RoboDK station: Senior Project 6612247056.rdk

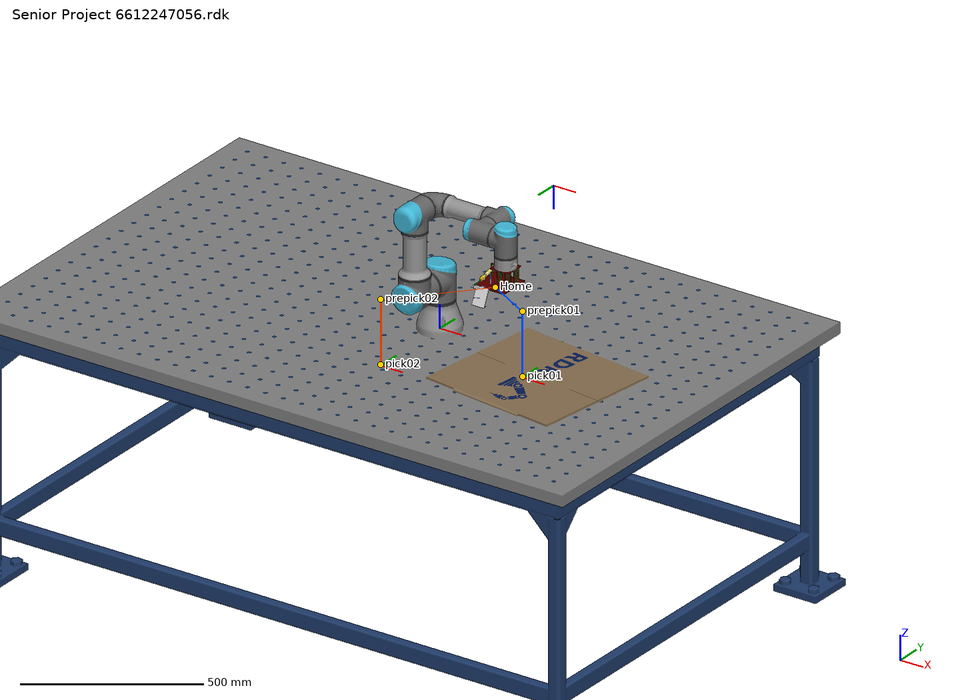
[picture v0: the station drawn from its stored meshes, robots at their saved joint values, targets as dots, program paths as lines]
Station Tast (saved by RoboDK 6.0.1). Poses are relative to the parent item; angles as X-Y-Z fixed-axis rotations.
  - frame Table at (0, 0, 0) mm
    - object Table at (-760, 0, 0) mm, size 2020 x 1340 x 800 mm, geometry from Table-2000x1200x800mm.sld
    - target Home (Cartesian target) at (261.4, -110.4, 243.15) mm, rotated rx -180 ry 0 rz -90 deg; joints [0, -90, -90, -90, 90, 0] of UR3
    - frame Camera 1 at (450, -100, 600) mm, rotated rx 180 ry 0 rz 0 deg
      - camera Camera 1
    - object BOX at (374.64, -51.63, 2) mm, rotated rx 0 ry 0.01 rz -7.34 deg, size 444 x 419.7 x 11.5 mm, geometry from Box-215x215mm-Unfolded.sld
  - frame UR3 Base at (0, 0, 0) mm
    - robot UR3: 6 axes, payload 3 kg, reach 500 mm, repeatability 0.1 mm, weight 11 kg
        modified DH rows (alpha deg, a mm, theta deg, d mm): 0, 0, 0, 151.9; 90, 0, 180, 0; 0, 243.65, 0, 0; 0, 213, 0, 110.4; -90, 0, 0, 83.4; 90, 0, 180, 82.4
        joint limits [-360, -360, -360, -360, -360, -360] to [360, 360, 360, 360, 360, 360]; home [0, -90, -90, 0, 90, 0]; saved at [0, -90, -90, -90, 90, 0]
      - tool Assem1, TCP at (0, 35, 70) mm, size 142.5 x 102 x 100.1 mm, geometry from Assem1.STEP
  - frame Orinal_Box at (360, -120, 0) mm
    - target prepick01 (Cartesian target) at (0, 0, 200) mm, rotated rx 180 ry 0 rz -90 deg; joints [20.517, -90.713, -100.969, -78.318, 90, 20.517] of UR3
    - target pick01 (Cartesian target) at (0, 0, 2) mm, rotated rx -180 ry 0 rz -90 deg; joints [-1.388, -136.982, -93.252, -39.765, 90.001, -1.388] of UR3
  - frame Orinal_Box(2) at (0, -280, 0) mm
    - target prepick02 (Cartesian target) at (0, 0, 200) mm, rotated rx -179.99 ry 0 rz 178.23 deg; joints [-68.924, -88.183, -103.474, -78.333, 90.001, 22.846] of UR3
    - target pick02 (Cartesian target) at (0, 0, 2) mm, rotated rx 179.99 ry 0 rz -179.49 deg; joints [-69.427, -124.075, -125.27, -20.665, 90, 20.063] of UR3
  - program Prog1 (1 instructions, listed below)
  - program pick (10 instructions, listed below)
  - program Place (8 instructions, listed below)
  - Python program Prog5 (listed below)
  - program Run (3 instructions, listed below)
  - Python program ur3_vision_pick_place (listed below)
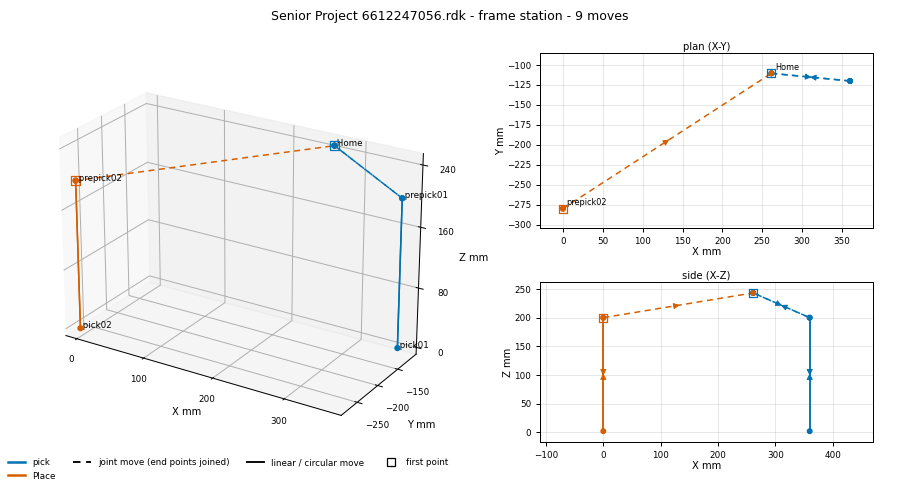
[picture p0: tool path of Senior Project 6612247056.rdk in frame station, 9 of 9 moves have a stored position in this frame; points joined in program order, loops and branches not executed]

--- program Prog1 (robot UR3) ---
  Move objects

--- program pick (robot UR3) ---
  ตั้งค่าRef: Table
  ตั้งค่าเครื่องมือ: Assem1
  MoveJ (Home)
  ตั้งค่าRef: Orinal_Box
  MoveJ (prepick01)
  MoveL (pick01)
  Attach to Assem1
  MoveL (prepick01)
  ตั้งค่าRef: Table
  MoveJ (Home)

--- program Place (robot UR3) ---
  ตั้งค่าRef: Orinal_Box(2)
  ตั้งค่าเครื่องมือ: Tool 1 at (0, 35, 70) mm
  MoveJ (prepick02)
  MoveL (pick02)
  ถอดออกจาก Assem1
  MoveL (prepick02)
  ตั้งค่าRef: Table
  MoveJ (Home)

--- Python program Prog5 ---
from robodk import robolink

RDK = robolink.Robolink()

# ดึงโปรแกรมมารันตรงๆ
prog_pick = RDK.Item('pick', robolink.ITEM_TYPE_PROGRAM)
prog_place = RDK.Item('Place', robolink.ITEM_TYPE_PROGRAM)

print("กำลังรันโปรแกรม Pick...")
prog_pick.RunProgram()


print("กำลังรันโปรแกรม Place...")
prog_place.RunProgram()

--- program Run (robot UR3) ---
  โทร Prog1
  โทร pick
  โทร Place

--- Python program ur3_vision_pick_place ---
"""
===============================================================================
UR3 Vision-Guided Pick & Place System with YOLOv8 & RoboDK
===============================================================================
Senior Project 6612247047
- YOLOv8 Model: Box_Logo.v2i.yolov8 (best (2).pt)
- RoboDK Station: Senior Project 6612247047 (UR3 Robot + Assem1 Gripper + BOX)
- Collision-Free Safe Execution via Home Posture
===============================================================================
"""

from robodk.robolink import *
from robodk.robomath import *
from ultralytics import YOLO
import cv2
import os
import time

# -----------------------------------------------------------------------------
# 1. Configuration & Initializations
# -----------------------------------------------------------------------------
MODEL_PATH = r'f:\New folder\best (2).pt'
SNAPSHOT_PATH = r'f:\New folder\temp_cam_snapshot.png'
ROBOT_SPEED = 80  # Speed in mm/s for safe motion

print("=" * 60)
print("  UR3 Vision-Guided Pick & Place System starting...")
print("=" * 60)

# Load YOLOv8 Model
if not os.path.exists(MODEL_PATH):
    raise FileNotFoundError(f"Model file not found at: {MODEL_PATH}")

print(f"[AI] Loading YOLOv8 model: {MODEL_PATH}...")
model = YOLO(MODEL_PATH)
print(f"[AI] Model classes loaded: {model.names}")

# Connect to RoboDK
print("[RoboDK] Connecting to RoboDK...")
RDK = Robolink()

if not RDK.Connect():
    print("[ERROR] Could not connect to RoboDK! Please ensure RoboDK is running.")
    exit(1)

station = RDK.ActiveStation()
print(f"[RoboDK] Connected to station: '{station.Name()}'")

# Get Items from RoboDK Station
robot = RDK.Item('UR3', ITEM_TYPE_ROBOT)
gripper = RDK.Item('Assem1', ITEM_TYPE_TOOL)
if not gripper.Valid():
    gripper = RDK.Item('gripper', ITEM_TYPE_TOOL)

target_item = RDK.Item('BOX', ITEM_TYPE_OBJECT)
if not target_item.Valid():
    target_item = RDK.Item('box', ITEM_TYPE_OBJECT)

home_target = RDK.Item('Home', ITEM_TYPE_TARGET)
prepick01 = RDK.Item('prepick01', ITEM_TYPE_TARGET)
pick01 = RDK.Item('pick01', ITEM_TYPE_TARGET)
prepick02 = RDK.Item('prepick02', ITEM_TYPE_TARGET)
pick02 = RDK.Item('pick02', ITEM_TYPE_TARGET)

table_frame = RDK.Item('Table', ITEM_TYPE_FRAME)
if not table_frame.Valid():
    table_frame = target_item.Parent()

cam_item = RDK.Item('Camera 1')

# Validate essential items
if not robot.Valid():
    print("[ERROR] Robot 'UR3' not found in RoboDK station!")
    exit(1)
if not target_item.Valid():
    print("[ERROR] Object 'BOX' not found in RoboDK station!")
    exit(1)

print("[RoboDK] All essential robot and station items loaded successfully.")

# Set safe robot speed
robot.setSpeed(ROBOT_SPEED)

# -----------------------------------------------------------------------------
# 2. Collision-Free Pick and Place Routine
# -----------------------------------------------------------------------------
def execute_safe_pick_and_place():
    """
    Executes a safe step-by-step pick and place operation for UR3:
    1. Move to Home (safe posture)
    2. Approach prepick01 (hover over source)
    3. Move to pick01 (pick position)
    4. Attach object BOX to gripper Assem1
    5. Retract up to prepick01
    6. Return to Home (safe transit posture avoiding self-collision)
    7. Move to prepick02 (hover over target destination)
    8. Move to pick02 (place position)
    9. Detach object BOX to table frame
    10. Retract up to prepick02
    11. Return safely to Home
    """
    print("\n" + "=" * 50)
    print(">>> STARTING COLLISION-FREE PICK & PLACE SEQUENCE <<<")
    print("=" * 50)

    # Step 1: Return to Home target (safe posture)
    print("Step 1/11: Moving to Home position...")
    if home_target.Valid():
        robot.setPoseFrame(home_target.Parent())
        robot.MoveJ(home_target)
    else:
        robot.MoveJ([0.0, -90.0, -90.0, -90.0, 90.0, 0.0])

    # Step 2: Move to prepick01 (hover above pick spot)
    print("Step 2/11: Approaching pick position (prepick01)...")
    if prepick01.Valid():
        robot.setPoseFrame(prepick01.Parent())
        robot.MoveJ(prepick01)

    # Step 3: Move down to pick01
    print("Step 3/11: Moving down to Pick (pick01)...")
    if pick01.Valid():
        robot.setPoseFrame(pick01.Parent())
        robot.MoveL(pick01)

    # Step 4: Attach object to gripper
    print("Step 4/11: Gripping / Attaching object 'BOX' to tool...")
    target_item.setParentStatic(gripper)
    time.sleep(0.5)

    # Step 5: Retract up to prepick01
    print("Step 5/11: Lifting object (prepick01)...")
    if prepick01.Valid():
        robot.setPoseFrame(prepick01.Parent())
        robot.MoveL(prepick01)

    # Step 6: Transit back to Home position (prevents arm rotation collision)
    print("Step 6/11: Returning to Home position for safe transit...")
    if home_target.Valid():
        robot.setPoseFrame(home_target.Parent())
        robot.MoveJ(home_target)

    # Step 7: Move to prepick02 (hover above place spot)
    print("Step 7/11: Approaching destination (prepick02)...")
    if prepick02.Valid():
        robot.setPoseFrame(prepick02.Parent())
        robot.MoveJ(prepick02)

    # Step 8: Move down to pick02 (place spot)
    print("Step 8/11: Moving down to Place (pick02)...")
    if pick02.Valid():
        robot.setPoseFrame(pick02.Parent())
        robot.MoveL(pick02)

    # Step 9: Detach object to Table frame
    print("Step 9/11: Releasing object 'BOX' onto target frame...")
    target_item.setParentStatic(table_frame)
    time.sleep(0.5)

    # Step 10: Retract up to prepick02
    print("Step 10/11: Retracting arm (prepick02)...")
    if prepick02.Valid():
        robot.setPoseFrame(prepick02.Parent())
        robot.MoveL(prepick02)

    # Step 11: Return to Home
    print("Step 11/11: Returning to Home position (Completed)...")
    if home_target.Valid():
        robot.setPoseFrame(home_target.Parent())
        robot.MoveJ(home_target)

    print("=" * 50)
    print(">>> PICK & PLACE COMPLETED SUCCESSFULLY WITH NO COLLISIONS <<<")
    print("=" * 50 + "\n")

# -----------------------------------------------------------------------------
# 3. Vision Loop (Webcam / RoboDK Camera Feed)
# -----------------------------------------------------------------------------
def run_vision_system():
    # Try opening webcam (index 0)
    cap = cv2.VideoCapture(0)
    use_robodk_cam = False

    if not cap.isOpened():
        print("[Camera] Physical webcam (index 0) not detected.")
        print("[Camera] Switching to RoboDK 'Camera 1' snapshot stream...")
        use_robodk_cam = True

    print("\nControls:")
    print(" - Press 'p' or 'SPACE' to trigger UR3 Pick & Place")
    print(" - Press 'q' to quit application")
    print("-" * 50)

    last_trigger_time = 0

    while True:
        frame = None

        if not use_robodk_cam:
            success, frame = cap.read()
            if not success:
                print("[Camera] Failed to grab frame from webcam. Switching to RoboDK camera...")
                use_robodk_cam = True

        if use_robodk_cam:
            if cam_item.Valid():
                RDK.Cam2D_Snapshot(SNAPSHOT_PATH, cam_item)
                if os.path.exists(SNAPSHOT_PATH):
                    frame = cv2.imread(SNAPSHOT_PATH)
            time.sleep(0.05)

        if frame is None:
            print("[Camera] Unable to capture frame!")
            time.sleep(0.5)
            continue

        # Run YOLOv8 detection
        results = model(frame, conf=0.25, verbose=False)
        annotated_frame = results[0].plot()

        box_detected = False
        detected_coords = []

        for r in results:
            for box in r.boxes:
                b = box.xyxy[0].cpu().numpy()
                cls_id = int(box.cls[0].item())
                cls_name = model.names.get(cls_id, str(cls_id))
                conf = float(box.conf[0].item())

                center_x = int((b[0] + b[2]) / 2)
                center_y = int((b[1] + b[3]) / 2)

                detected_coords.append((cls_name, center_x, center_y, conf))
                box_detected = True

                # Draw center point and coordinates text
                cv2.circle(annotated_frame, (center_x, center_y), 5, (0, 255, 0), -1)
                cv2.putText(
                    annotated_frame,
                    f"{cls_name} ({center_x},{center_y})",
                    (center_x - 40, center_y - 10),
                    cv2.FONT_HERSHEY_SIMPLEX,
                    0.5,
                    (0, 255, 0),
                    2
                )

        # Status text overlay
        cam_type_str = "RoboDK Camera 1" if use_robodk_cam else "Webcam (0)"
        cv2.putText(
            annotated_frame,
            f"Cam: {cam_type_str} | Press 'p' to Pick&Place | 'q' to Quit",
            (10, 30),
            cv2.FONT_HERSHEY_SIMPLEX,
            0.6,
            (255, 255, 0),
            2
        )

        # Display OpenCV Window
        cv2.imshow("Senior Project 6612247047 - UR3 Vision System (YOLOv8)", annotated_frame)

        key = cv2.waitKey(1) & 0xFF
        if key == ord('q'):
            print("[System] User requested exit.")
            break
        elif key in (ord('p'), ord(' '), ord('P')):
            # Trigger pick & place operation
            current_time = time.time()
            if current_time - last_trigger_time > 3.0:
                print(f"\n[Trigger] Pick & Place triggered! Detected objects: {detected_coords}")
                execute_safe_pick_and_place()
                last_trigger_time = time.time()

    if not use_robodk_cam and cap:
        cap.release()
    cv2.destroyAllWindows()
    print("[System] Vision system shut down successfully.")

# -----------------------------------------------------------------------------
# Main Entry Point
# -----------------------------------------------------------------------------
if __name__ == "__main__":
    run_vision_system()
